FUNCTION_BLOCK FB_LivingRoom
VAR
    // Logical input placeholders. Map these to physical terminals later.
    bCeilingSwitchInput : BOOL;
    bWallSwitchInput    : BOOL;
    bAmbientSwitchInput : BOOL;

    stCeilingSwitchId : ST_DeviceId;
    stWallSwitchId    : ST_DeviceId;
    stAmbientSwitchId : ST_DeviceId;

    fbCeilingSwitch : FB_SwitchMonostable;
    fbWallSwitch    : FB_SwitchMonostable;
    fbAmbientSwitch : FB_SwitchMonostable;

    fbCeilingSwitchCtrl : FB_SwitchCtrl;
    fbWallSwitchCtrl    : FB_SwitchCtrl;
    fbAmbientSwitchCtrl : FB_SwitchCtrl;
END_VAR

stCeilingSwitchId.sId := 101;
stCeilingSwitchId.sName := 'Ceiling Switch';
stCeilingSwitchId.sRoom := 'Living Room';

stWallSwitchId.sId := 102;
stWallSwitchId.sName := 'Wall Switch';
stWallSwitchId.sRoom := 'Living Room';

stAmbientSwitchId.sId := 103;
stAmbientSwitchId.sName := 'Ambient Switch';
stAmbientSwitchId.sRoom := 'Living Room';

fbCeilingSwitch(stDeviceId := stCeilingSwitchId, bInput := bCeilingSwitchInput);
fbWallSwitch(stDeviceId := stWallSwitchId, bInput := bWallSwitchInput);
fbAmbientSwitch(stDeviceId := stAmbientSwitchId, bInput := bAmbientSwitchInput);

fbCeilingSwitchCtrl(iSwitch := fbCeilingSwitch);
fbWallSwitchCtrl(iSwitch := fbWallSwitch);
fbAmbientSwitchCtrl(iSwitch := fbAmbientSwitch);

// Room logic writes commands; FB_House resets command pulses once per scan.
IF fbCeilingSwitchCtrl.stControlData.bShortClick THEN
    CASE fbCeilingSwitchCtrl.stControlData.nShortClickCount OF
        1:
            GVL_LightCmds.stLivingRoomCeilingCmd.eAction := E_LightAction.Toggle;
        2:
            GVL_LightCmds.stLivingRoomCeilingCmd.eAction := E_LightAction.SetBrightness;
            GVL_LightCmds.stLivingRoomCeilingCmd.nBrightness := 40;
        4:
            GVL_LightCmds.stLivingRoomCeilingCmd.eAction := E_LightAction.TurnOff;
            GVL_LightCmds.stLivingRoomWallCmd.eAction := E_LightAction.TurnOff;
            GVL_LightCmds.stLivingRoomAmbientCmd.eAction := E_LightAction.TurnOff;
    END_CASE
END_IF

IF fbWallSwitchCtrl.stControlData.bShortClick AND
   (fbWallSwitchCtrl.stControlData.nShortClickCount = 1) THEN
    GVL_LightCmds.stLivingRoomWallCmd.eAction := E_LightAction.Toggle;
END_IF

IF fbAmbientSwitchCtrl.stControlData.bShortClick AND
   (fbAmbientSwitchCtrl.stControlData.nShortClickCount = 1) THEN
    GVL_LightCmds.stLivingRoomAmbientCmd.eAction := E_LightAction.Toggle;
END_IF

END_FUNCTION_BLOCK

(* stored: Version 1.1.0.1, ProductVersion 3.1.4026.20
   POU FB_LivingRoom: Id {D4E8A210-3B71-4C96-8F25-7A1B2C3D4001} *)
